PROGRAM main
  VAR
    B1 AT %IX0.0     : BOOL; (* sensor de cajas *)
    KM1 AT %QX0.0    : BOOL; (* banda (bobina 00001 para la PC) *)
    CAJAS AT %MW0    : INT; (* holding 40001: cajas contadas *)
    P_MARCHA AT %MW1 : INT; (* holding 40002: pulsador remoto MARCHA *)
    P_PARO AT %MW2   : INT; (* holding 40003: pulsador remoto PARO *)
    P_CERO AT %MW3   : INT; (* holding 40004: pulsador remoto contador a cero *)
    F_CAJA           : R_TRIG;
    CAJA             : BOOL; (* flanco de B1 *)
  END_VAR
  VAR  (* added by the conversion: wires and edge detectors of the diagram *)
    _NE5_OUT : BOOL;
    _ADD11_OUT : INT;
    _SEL8_OUT : INT;
    _SEL4_OUT : INT;
    _NE19_OUT : BOOL;
    _OR17_OUT : BOOL;
    _EQ22_OUT : BOOL;
    _AND16_OUT : BOOL;
    _NE27_OUT : BOOL;
    _SEL26_OUT : INT;
    _NE34_OUT : BOOL;
    _SEL33_OUT : INT;
    _NE41_OUT : BOOL;
    _SEL40_OUT : INT;
  END_VAR

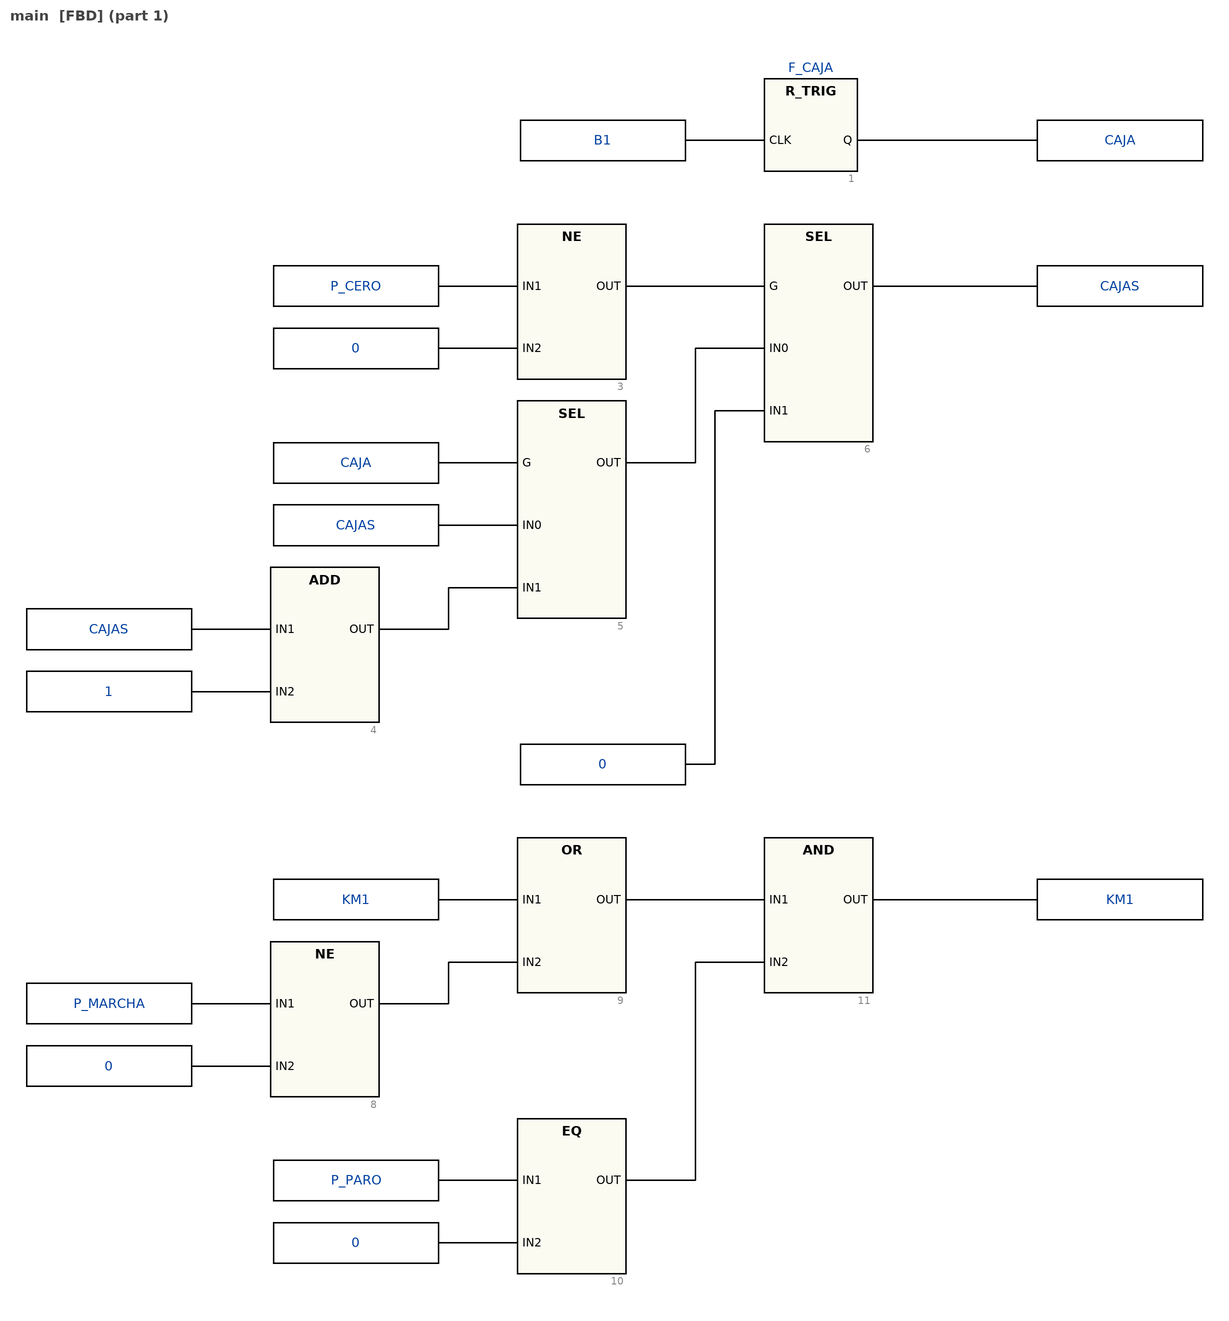
(* FBD diagram, written out as Structured Text *)
F_CAJA(CLK := B1);
CAJA := F_CAJA.Q;
_NE5_OUT := P_CERO <> 0;
_ADD11_OUT := CAJAS + 1;
_SEL8_OUT := SEL(CAJA, CAJAS, _ADD11_OUT);
_SEL4_OUT := SEL(_NE5_OUT, _SEL8_OUT, 0);
CAJAS := _SEL4_OUT;
_NE19_OUT := P_MARCHA <> 0;
_OR17_OUT := KM1 OR _NE19_OUT;
_EQ22_OUT := P_PARO = 0;
_AND16_OUT := _OR17_OUT AND _EQ22_OUT;
KM1 := _AND16_OUT;
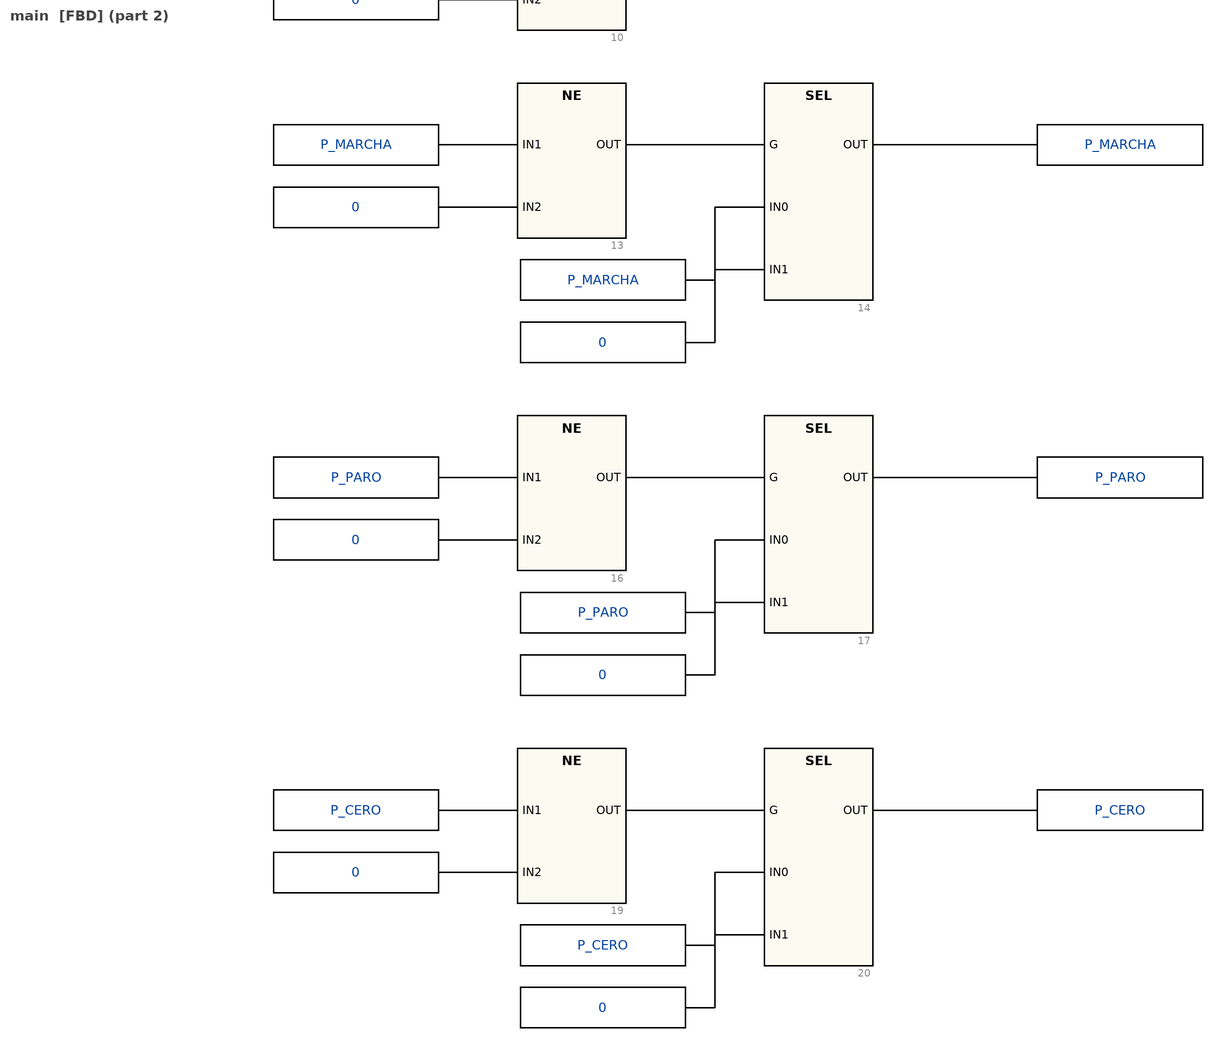
_NE27_OUT := P_MARCHA <> 0;
_SEL26_OUT := SEL(_NE27_OUT, P_MARCHA, 0);
P_MARCHA := _SEL26_OUT;
_NE34_OUT := P_PARO <> 0;
_SEL33_OUT := SEL(_NE34_OUT, P_PARO, 0);
P_PARO := _SEL33_OUT;
_NE41_OUT := P_CERO <> 0;
_SEL40_OUT := SEL(_NE41_OUT, P_CERO, 0);
P_CERO := _SEL40_OUT;
END_PROGRAM
